// TIA Portal V20 export
FUNCTION_BLOCK "PR_StackUltraWeldSeq_Soft2"   // FB55, LAD
{ S7_Optimized_Access := 'TRUE' }
// stored: MemoryReserve 100, SetENOAutomatically false
   VAR_INPUT
      iAbort : Bool;
      iAutoRunning : Bool;
      iFaultReset : Bool;
      iPartClampClose : Bool;
      iPartClampOpen : Bool;
      iPartNotWorkable : Bool;
      iPartWorkable : Bool;
      iRFReadDone : Bool;
      iRFReadError : Bool;
      iRFWriteDone : Bool;
      iRFWriteError : Bool;
      iReject : Bool;
      iReset_fault : Bool;
      iRetry : Bool;
      iRetryCount : Int;
      iSstMode : Bool;
      iSstPB : Bool;
      iStartFrmFibroseq : Bool;
      iWeldComplete : Bool;
      iWeldTabDown : Bool;
      iWeldTabUp : Bool;
      iStartFrmFibroSeq_1 : Bool;
      iAutorunning_1 : Bool;
   END_VAR
   VAR_OUTPUT
      qError : Array[0..3] of Bool;
      qFumeExtractorON : Bool;
      qMessage : Array[0..2] of Bool;
      qPartClampClose : Bool;
      qPartClampOpen : Bool;
      qStackUltraWeldOver : Bool;
      qWeldTabDown : Bool;
      qWeldTabUp : Bool;
   END_VAR
   VAR
      c20_ChkRecovery_T1 : Bool;
      c20_ChkRecovery_T2 : Bool;
      c20_ChkRecovery_T3 : Bool;
      c21_WtRFIDReadOver_T1 : Bool;
      c21_WtRFIDReadOver_T2 : Bool;
      c22_ChkReadRetryCnt_T1 : Bool;
      c22_ChkReadRetryCnt_T2 : Bool;
      c23_ChkPartWrkSts_T1 : Bool;
      c23_ChkPartWrkSts_T2 : Bool;
      c24_WtOpDecision_T1 : Bool;
      c24_WtOpDecision_T2 : Bool;
      c81_WtRFIDWriteOver_T1 : Bool;
      c81_WtRFIDWriteOver_T2 : Bool;
      c82_ChkWriteRetryCnt_T1 : Bool;
      c82_ChkWriteRetryCnt_T2 : Bool;
      c83_WtOpDecisionWrite_T1 : Bool;
      c83_WtOpDecisionWrite_T2 : Bool;
      StateNo : Int;
      s10_WtStartFrmFibro : Bool;
      s10_WtStartFrmFibro_T1 : Bool;
      s1_WtResetRel : Bool;
      s1_WtResetRel_T1 : Bool;
      s20_ChkRecovery : Bool;
      s20_ChkRecovery_T1 : Bool;
      s20_ChkRecovery_T2 : Bool;
      s20_ChkRecovery_T3 : Bool;
      s21_WtRFIDReadOver : Bool;
      s21_WtRFIDReadOver_T1 : Bool;
      s21_WtRFIDReadOver_T2 : Bool;
      s22_ChkReadRetryCnt : Bool;
      s22_ChkReadRetryCnt_T1 : Bool;
      s22_ChkReadRetryCnt_T2 : Bool;
      s23_ChkPartWrkSts : Bool;
      s23_ChkPartWrkSts_T1 : Bool;
      s23_ChkPartWrkSts_T2 : Bool;
      s24_WtOpDecision : Bool;
      s24_WtOpDecision_T1 : Bool;
      s24_WtOpDecision_T2 : Bool;
      s30_WtOpAck : Bool;
      s30_WtOpAck_T1 : Bool;
      s40_WtPartClamp : Bool;
      s40_WtPartClamp_T1 : Bool;
      s50_WtWeldTabDown : Bool;
      s50_WtWeldTabDown_T1 : Bool;
      s60_WtWeldComplete : Bool;
      s60_WtWeldComplete_T1 : Bool;
      s70_WtWeldTabUp : Bool;
      s70_WtWeldTabUp_T1 : Bool;
      s80_WtPartClampOpen : Bool;
      s80_WtPartClampOpen_T1 : Bool;
      s81_WtRFIDWriteOver : Bool;
      s81_WtRFIDWriteOver_T1 : Bool;
      s81_WtRFIDWriteOver_T2 : Bool;
      s82_ChkWriteRetryCnt : Bool;
      s82_ChkWriteRetryCnt_T1 : Bool;
      s82_ChkWriteRetryCnt_T2 : Bool;
      s83_WtOpDecisionWrite : Bool;
      s83_WtOpDecisionWrite_T1 : Bool;
      s83_WtOpDecisionWrite_T2 : Bool;
      s90_WtStartLow : Bool;
      s90_WtStartLow_T1 : Bool;
      sRFReadRetryCount : Int;
      sRFWriteRetryCount : Int;
      sSst : Bool;
      sSstPulse : Bool;
      sSstRise : Bool;
      sStWtResetRel : Bool;
      sStWtResetRel_T1 : Bool;
      sWeldDlyOver : Bool;
      sweldingInProgress : Int;
      SET : Bool;
      c20_ChkRecovery_clamp : Bool;
   END_VAR
   VAR_TEMP
      tOne : Bool;
      tRFReadRetryCountInc : Int;
      tRFWriteRetryCountInc : Int;
   END_VAR
   VAR_TEMP   // added for the SCL form of the ladder/FBD networks
      _w1 : Bool;
      _w2 : Bool;
   END_VAR
BEGIN

REGION Network 1
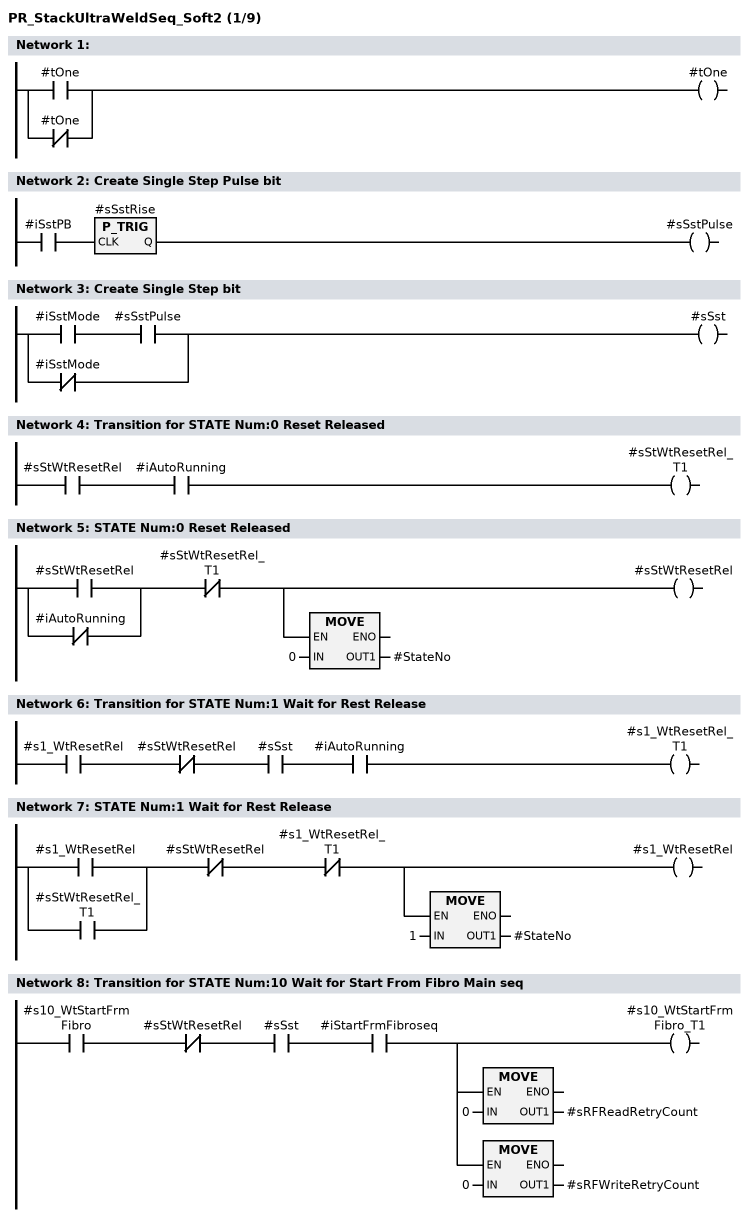
   RUNG wire#powerrail
      Contact( #tOne )
      wire#w1
      Coil( #tOne )
   END_RUNG
   RUNG wire#powerrail
      I_Contact( #tOne )
   END_RUNG wire#w1
   // the same network as SCL:
   #tOne := #tOne OR NOT #tOne;
END_REGION

REGION Network 2: Create Single Step Pulse bit
   RUNG wire#powerrail
      Contact( #iSstPB )
      P_Trig( #sSstRise )
      Coil( #sSstPulse )
   END_RUNG
   // the same network as SCL:
   #_w1 := #iSstPB AND NOT #sSstRise;   // rising edge
   #sSstRise := #iSstPB;
   #sSstPulse := #_w1;
END_REGION

REGION Network 3: Create Single Step bit
   RUNG wire#powerrail
      Contact( #iSstMode )
      Contact( #sSstPulse )
      wire#w1
      Coil( #sSst )
   END_RUNG
   RUNG wire#powerrail
      I_Contact( #iSstMode )
   END_RUNG wire#w1
   // the same network as SCL:
   #sSst := (#iSstMode AND #sSstPulse) OR NOT #iSstMode;
END_REGION

REGION Network 4: Transition for STATE Num:0 Reset Released
   RUNG wire#powerrail
      Contact( #sStWtResetRel )
      Contact( #iAutoRunning )
      Coil( #sStWtResetRel_T1 )
   END_RUNG
   // the same network as SCL:
   #sStWtResetRel_T1 := #sStWtResetRel AND #iAutoRunning;
END_REGION

REGION Network 5: STATE Num:0 Reset Released
   RUNG wire#powerrail
      Contact( #sStWtResetRel )
      wire#w1
      I_Contact( #sStWtResetRel_T1 )
      wire#w2
      Coil( #sStWtResetRel )
   END_RUNG
   RUNG wire#powerrail
      I_Contact( #iAutoRunning )
   END_RUNG wire#w1
   RUNG wire#w2
      { S7_GenerateENO := "TRUE" } Move(in := 0, out1 => #StateNo)
   END_RUNG
   // the same network as SCL:
   #sStWtResetRel := (#sStWtResetRel OR NOT #iAutoRunning) AND NOT #sStWtResetRel_T1;
   IF #sStWtResetRel THEN #StateNo := 0; END_IF;
END_REGION

REGION Network 6: Transition for STATE Num:1 Wait for Rest Release
   RUNG wire#powerrail
      Contact( #s1_WtResetRel )
      I_Contact( #sStWtResetRel )
      Contact( #sSst )
      Contact( #iAutoRunning )
      Coil( #s1_WtResetRel_T1 )
   END_RUNG
   // the same network as SCL:
   #s1_WtResetRel_T1 := #s1_WtResetRel AND NOT #sStWtResetRel AND #sSst AND #iAutoRunning;
END_REGION

REGION Network 7: STATE Num:1 Wait for Rest Release
   RUNG wire#powerrail
      Contact( #s1_WtResetRel )
      wire#w1
      I_Contact( #sStWtResetRel )
      I_Contact( #s1_WtResetRel_T1 )
      wire#w2
      Coil( #s1_WtResetRel )
   END_RUNG
   RUNG wire#powerrail
      Contact( #sStWtResetRel_T1 )
   END_RUNG wire#w1
   RUNG wire#w2
      { S7_GenerateENO := "TRUE" } Move(in := 1, out1 => #StateNo)
   END_RUNG
   // the same network as SCL:
   #s1_WtResetRel := (#s1_WtResetRel OR #sStWtResetRel_T1) AND NOT #sStWtResetRel AND NOT #s1_WtResetRel_T1;
   IF #s1_WtResetRel THEN #StateNo := 1; END_IF;
END_REGION

REGION Network 8: Transition for STATE Num:10 Wait for Start From Fibro Main seq
   RUNG wire#powerrail
      Contact( #s10_WtStartFrmFibro )
      I_Contact( #sStWtResetRel )
      Contact( #sSst )
      Contact( #iStartFrmFibroseq )
      wire#w1
      Coil( #s10_WtStartFrmFibro_T1 )
   END_RUNG
   RUNG wire#w1
      Move(in := 0, out1 => #sRFReadRetryCount)
   END_RUNG
   RUNG wire#w1
      Move(in := 0, out1 => #sRFWriteRetryCount)
   END_RUNG
   // the same network as SCL:
   #s10_WtStartFrmFibro_T1 := #s10_WtStartFrmFibro AND NOT #sStWtResetRel AND #sSst AND #iStartFrmFibroseq;
   IF #s10_WtStartFrmFibro_T1 THEN
       #sRFReadRetryCount := 0;
       #sRFWriteRetryCount := 0;
   END_IF;
END_REGION

REGION Network 9: STATE Num:10 Wait for Start From Fibro Main seq
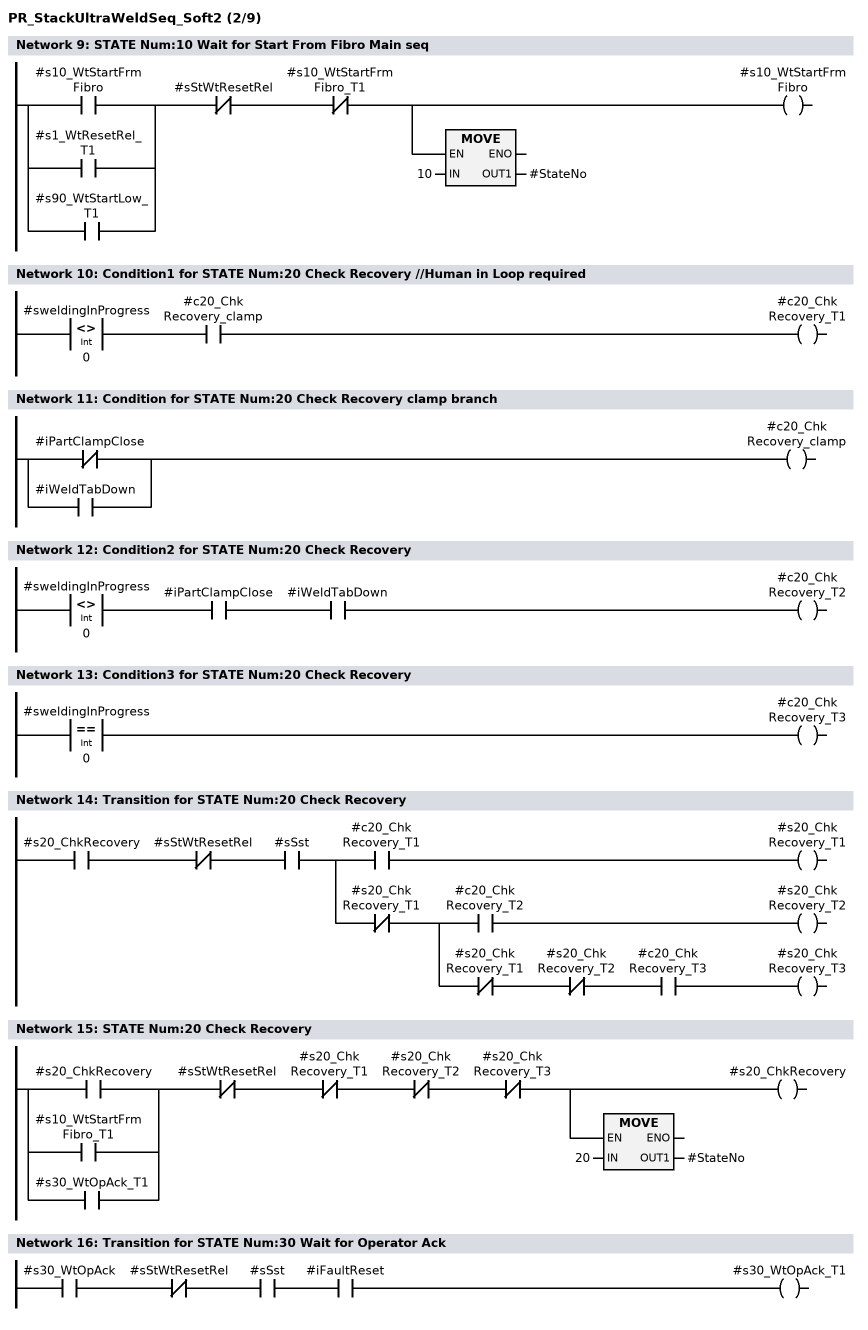
   RUNG wire#powerrail
      Contact( #s10_WtStartFrmFibro )
      wire#w1
      I_Contact( #sStWtResetRel )
      I_Contact( #s10_WtStartFrmFibro_T1 )
      wire#w2
      Coil( #s10_WtStartFrmFibro )
   END_RUNG
   RUNG wire#powerrail
      Contact( #s1_WtResetRel_T1 )
   END_RUNG wire#w1
   RUNG wire#powerrail
      Contact( #s90_WtStartLow_T1 )
   END_RUNG wire#w1
   RUNG wire#w2
      { S7_GenerateENO := "TRUE" } Move(in := 10, out1 => #StateNo)
   END_RUNG
   // the same network as SCL:
   #s10_WtStartFrmFibro := (#s10_WtStartFrmFibro OR #s1_WtResetRel_T1 OR #s90_WtStartLow_T1) AND NOT #sStWtResetRel AND NOT #s10_WtStartFrmFibro_T1;
   IF #s10_WtStartFrmFibro THEN #StateNo := 10; END_IF;
END_REGION

REGION Network 10: Condition1 for STATE Num:20 Check Recovery //Human in Loop required
   RUNG wire#powerrail
      { S7_Templates := "SrcType := Int" } NE_Contact(in1 := #sweldingInProgress, in2 := 0)
      Contact( #c20_ChkRecovery_clamp )
      Coil( #c20_ChkRecovery_T1 )
   END_RUNG
   // the same network as SCL:
   #c20_ChkRecovery_T1 := (#sweldingInProgress <> 0) AND #c20_ChkRecovery_clamp;
END_REGION

REGION Network 11: Condition for STATE Num:20 Check Recovery clamp branch
   RUNG wire#powerrail
      I_Contact( #iPartClampClose )
      wire#w1
      Coil( #c20_ChkRecovery_clamp )
   END_RUNG
   RUNG wire#powerrail
      Contact( #iWeldTabDown )
   END_RUNG wire#w1
   // the same network as SCL:
   #c20_ChkRecovery_clamp := NOT #iPartClampClose OR #iWeldTabDown;
END_REGION

REGION Network 12: Condition2 for STATE Num:20 Check Recovery
   RUNG wire#powerrail
      { S7_Templates := "SrcType := Int" } NE_Contact(in1 := #sweldingInProgress, in2 := 0)
      Contact( #iPartClampClose )
      Contact( #iWeldTabDown )
      Coil( #c20_ChkRecovery_T2 )
   END_RUNG
   // the same network as SCL:
   #c20_ChkRecovery_T2 := (#sweldingInProgress <> 0) AND #iPartClampClose AND #iWeldTabDown;
END_REGION

REGION Network 13: Condition3 for STATE Num:20 Check Recovery
   RUNG wire#powerrail
      { S7_Templates := "SrcType := Int" } EQ_Contact(in1 := #sweldingInProgress, in2 := 0)
      Coil( #c20_ChkRecovery_T3 )
   END_RUNG
   // the same network as SCL:
   #c20_ChkRecovery_T3 := #sweldingInProgress = 0;
END_REGION

REGION Network 14: Transition for STATE Num:20 Check Recovery
   RUNG wire#powerrail
      Contact( #s20_ChkRecovery )
      I_Contact( #sStWtResetRel )
      Contact( #sSst )
      wire#w1
      Contact( #c20_ChkRecovery_T1 )
      Coil( #s20_ChkRecovery_T1 )
   END_RUNG
   RUNG wire#w1
      I_Contact( #s20_ChkRecovery_T1 )
      wire#w2
      Contact( #c20_ChkRecovery_T2 )
      Coil( #s20_ChkRecovery_T2 )
   END_RUNG
   RUNG wire#w2
      I_Contact( #s20_ChkRecovery_T1 )
      I_Contact( #s20_ChkRecovery_T2 )
      Contact( #c20_ChkRecovery_T3 )
      Coil( #s20_ChkRecovery_T3 )
   END_RUNG
   // the same network as SCL:
   #_w1 := #s20_ChkRecovery AND NOT #sStWtResetRel AND #sSst;
   #s20_ChkRecovery_T1 := #_w1 AND #c20_ChkRecovery_T1;
   #_w2 := #_w1 AND NOT #s20_ChkRecovery_T1;
   #s20_ChkRecovery_T2 := #_w2 AND #c20_ChkRecovery_T2;
   #s20_ChkRecovery_T3 := #_w2 AND NOT #s20_ChkRecovery_T1 AND NOT #s20_ChkRecovery_T2 AND #c20_ChkRecovery_T3;
END_REGION

REGION Network 15: STATE Num:20 Check Recovery
   RUNG wire#powerrail
      Contact( #s20_ChkRecovery )
      wire#w1
      I_Contact( #sStWtResetRel )
      I_Contact( #s20_ChkRecovery_T1 )
      I_Contact( #s20_ChkRecovery_T2 )
      I_Contact( #s20_ChkRecovery_T3 )
      wire#w2
      Coil( #s20_ChkRecovery )
   END_RUNG
   RUNG wire#powerrail
      Contact( #s10_WtStartFrmFibro_T1 )
   END_RUNG wire#w1
   RUNG wire#powerrail
      Contact( #s30_WtOpAck_T1 )
   END_RUNG wire#w1
   RUNG wire#w2
      { S7_GenerateENO := "TRUE" } Move(in := 20, out1 => #StateNo)
   END_RUNG
   // the same network as SCL:
   #s20_ChkRecovery := (#s20_ChkRecovery OR #s10_WtStartFrmFibro_T1 OR #s30_WtOpAck_T1) AND NOT #sStWtResetRel AND NOT #s20_ChkRecovery_T1 AND NOT #s20_ChkRecovery_T2 AND NOT #s20_ChkRecovery_T3;
   IF #s20_ChkRecovery THEN #StateNo := 20; END_IF;
END_REGION

REGION Network 16: Transition for STATE Num:30 Wait for Operator Ack
   RUNG wire#powerrail
      Contact( #s30_WtOpAck )
      I_Contact( #sStWtResetRel )
      Contact( #sSst )
      Contact( #iFaultReset )
      Coil( #s30_WtOpAck_T1 )
   END_RUNG
   // the same network as SCL:
   #s30_WtOpAck_T1 := #s30_WtOpAck AND NOT #sStWtResetRel AND #sSst AND #iFaultReset;
END_REGION

REGION Network 17: STATE Num:30 Wait for Operator Ack
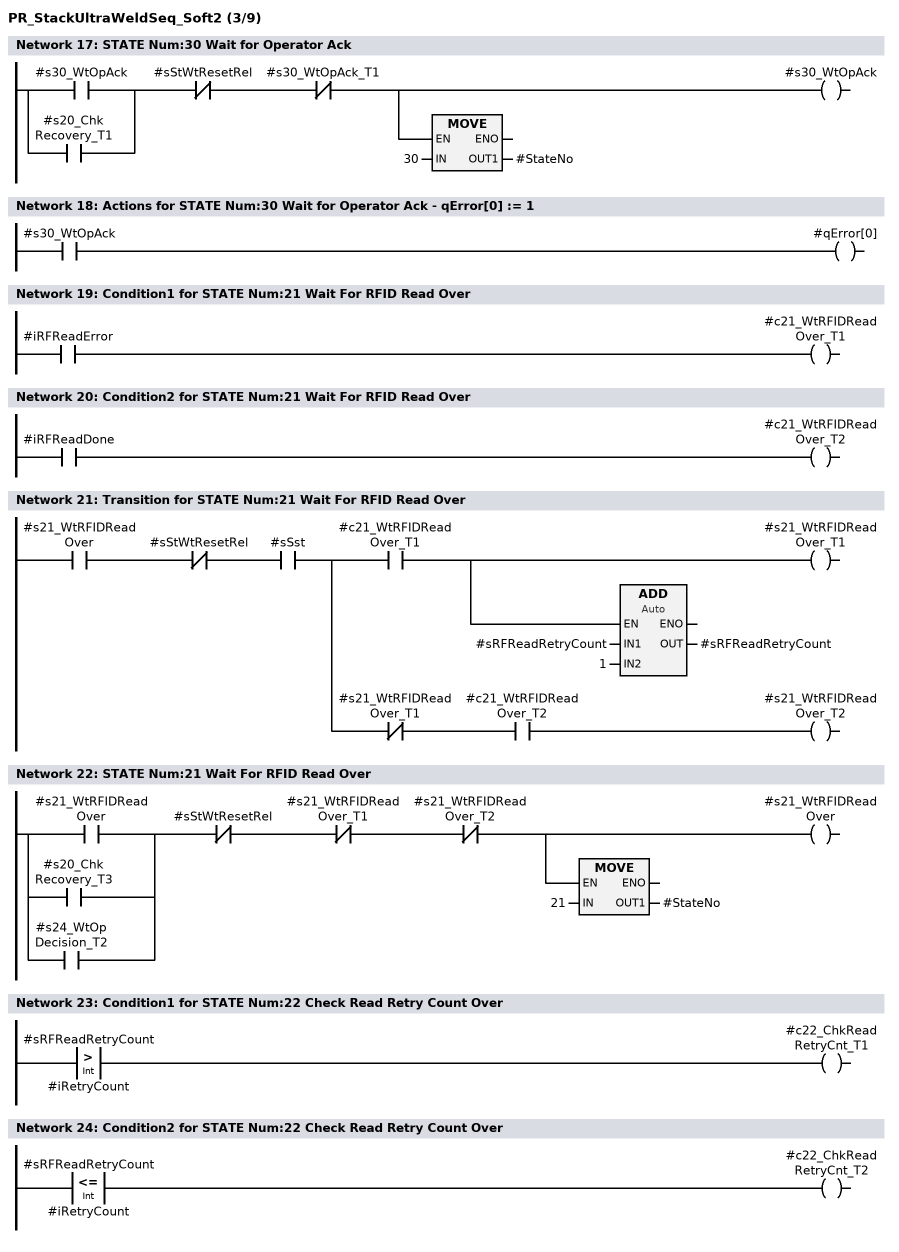
   RUNG wire#powerrail
      Contact( #s30_WtOpAck )
      wire#w1
      I_Contact( #sStWtResetRel )
      I_Contact( #s30_WtOpAck_T1 )
      wire#w2
      Coil( #s30_WtOpAck )
   END_RUNG
   RUNG wire#powerrail
      Contact( #s20_ChkRecovery_T1 )
   END_RUNG wire#w1
   RUNG wire#w2
      { S7_GenerateENO := "TRUE" } Move(in := 30, out1 => #StateNo)
   END_RUNG
   // the same network as SCL:
   #s30_WtOpAck := (#s30_WtOpAck OR #s20_ChkRecovery_T1) AND NOT #sStWtResetRel AND NOT #s30_WtOpAck_T1;
   IF #s30_WtOpAck THEN #StateNo := 30; END_IF;
END_REGION

REGION Network 18: Actions for STATE Num:30 Wait for Operator Ack - qError[0] := 1
   RUNG wire#powerrail
      Contact( #s30_WtOpAck )
      Coil( #qError[0] )
   END_RUNG
   // the same network as SCL:
   #qError[0] := #s30_WtOpAck;
END_REGION

REGION Network 19: Condition1 for STATE Num:21 Wait For RFID Read Over
   RUNG wire#powerrail
      Contact( #iRFReadError )
      Coil( #c21_WtRFIDReadOver_T1 )
   END_RUNG
   // the same network as SCL:
   #c21_WtRFIDReadOver_T1 := #iRFReadError;
END_REGION

REGION Network 20: Condition2 for STATE Num:21 Wait For RFID Read Over
   RUNG wire#powerrail
      Contact( #iRFReadDone )
      Coil( #c21_WtRFIDReadOver_T2 )
   END_RUNG
   // the same network as SCL:
   #c21_WtRFIDReadOver_T2 := #iRFReadDone;
END_REGION

REGION Network 21: Transition for STATE Num:21 Wait For RFID Read Over
   RUNG wire#powerrail
      Contact( #s21_WtRFIDReadOver )
      I_Contact( #sStWtResetRel )
      Contact( #sSst )
      wire#w1
      Contact( #c21_WtRFIDReadOver_T1 )
      wire#w2
      Coil( #s21_WtRFIDReadOver_T1 )
   END_RUNG
   RUNG wire#w2
      Add(in1 := #sRFReadRetryCount, in2 := 1, out => #sRFReadRetryCount)
   END_RUNG
   RUNG wire#w1
      I_Contact( #s21_WtRFIDReadOver_T1 )
      Contact( #c21_WtRFIDReadOver_T2 )
      Coil( #s21_WtRFIDReadOver_T2 )
   END_RUNG
   // the same network as SCL:
   #_w1 := #s21_WtRFIDReadOver AND NOT #sStWtResetRel AND #sSst;
   #s21_WtRFIDReadOver_T1 := #_w1 AND #c21_WtRFIDReadOver_T1;
   IF #s21_WtRFIDReadOver_T1 THEN #sRFReadRetryCount := #sRFReadRetryCount + 1; END_IF;
   #s21_WtRFIDReadOver_T2 := #_w1 AND NOT #s21_WtRFIDReadOver_T1 AND #c21_WtRFIDReadOver_T2;
END_REGION

REGION Network 22: STATE Num:21 Wait For RFID Read Over
   RUNG wire#powerrail
      Contact( #s21_WtRFIDReadOver )
      wire#w1
      I_Contact( #sStWtResetRel )
      I_Contact( #s21_WtRFIDReadOver_T1 )
      I_Contact( #s21_WtRFIDReadOver_T2 )
      wire#w2
      Coil( #s21_WtRFIDReadOver )
   END_RUNG
   RUNG wire#powerrail
      Contact( #s20_ChkRecovery_T3 )
   END_RUNG wire#w1
   RUNG wire#powerrail
      Contact( #s24_WtOpDecision_T2 )
   END_RUNG wire#w1
   RUNG wire#w2
      { S7_GenerateENO := "TRUE" } Move(in := 21, out1 => #StateNo)
   END_RUNG
   // the same network as SCL:
   #s21_WtRFIDReadOver := (#s21_WtRFIDReadOver OR #s20_ChkRecovery_T3 OR #s24_WtOpDecision_T2) AND NOT #sStWtResetRel AND NOT #s21_WtRFIDReadOver_T1 AND NOT #s21_WtRFIDReadOver_T2;
   IF #s21_WtRFIDReadOver THEN #StateNo := 21; END_IF;
END_REGION

REGION Network 23: Condition1 for STATE Num:22 Check Read Retry Count Over
   RUNG wire#powerrail
      { S7_Templates := "SrcType := Int" } GT_Contact(in1 := #sRFReadRetryCount, in2 := #iRetryCount)
      Coil( #c22_ChkReadRetryCnt_T1 )
   END_RUNG
   // the same network as SCL:
   #c22_ChkReadRetryCnt_T1 := #sRFReadRetryCount > #iRetryCount;
END_REGION

REGION Network 24: Condition2 for STATE Num:22 Check Read Retry Count Over
   RUNG wire#powerrail
      { S7_Templates := "SrcType := Int" } LE_Contact(in1 := #sRFReadRetryCount, in2 := #iRetryCount)
      Coil( #c22_ChkReadRetryCnt_T2 )
   END_RUNG
   // the same network as SCL:
   #c22_ChkReadRetryCnt_T2 := #sRFReadRetryCount <= #iRetryCount;
END_REGION

REGION Network 25: Transition for STATE Num:22 Check Read Retry Count Over
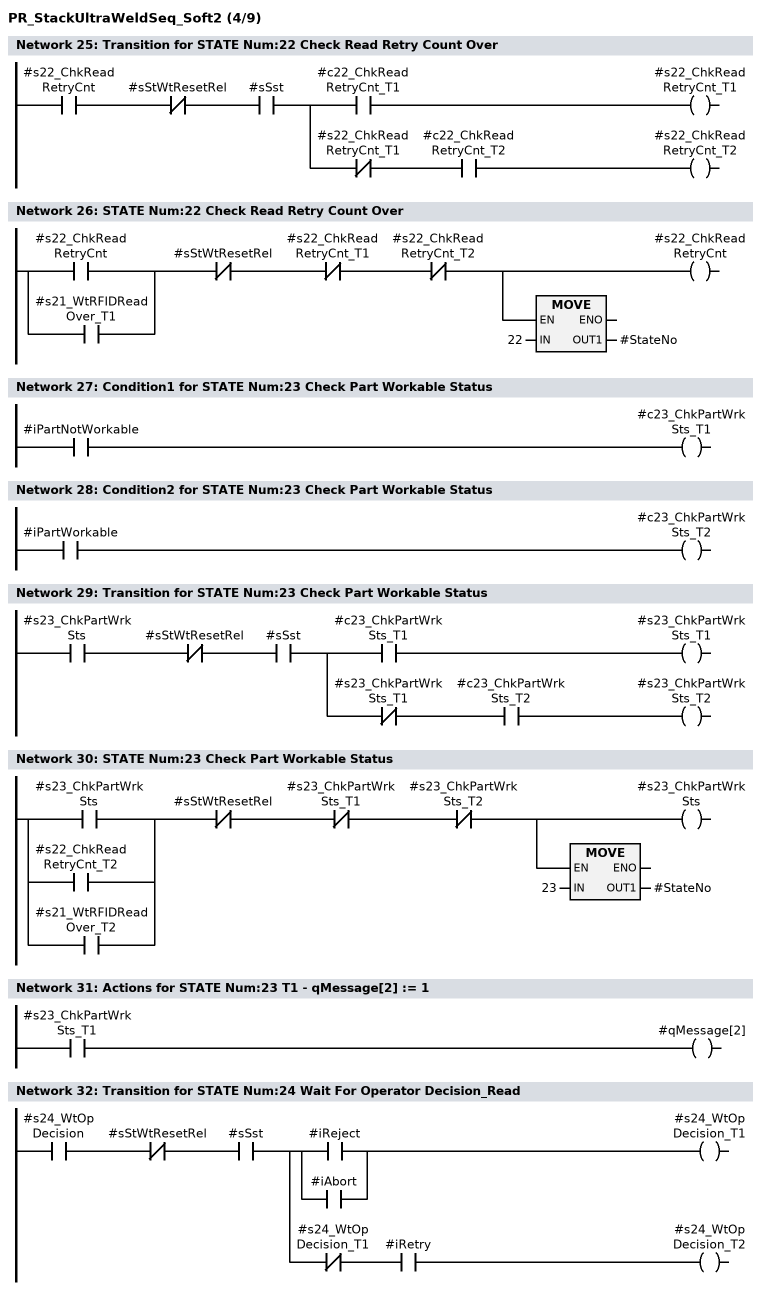
   RUNG wire#powerrail
      Contact( #s22_ChkReadRetryCnt )
      I_Contact( #sStWtResetRel )
      Contact( #sSst )
      wire#w1
      Contact( #c22_ChkReadRetryCnt_T1 )
      Coil( #s22_ChkReadRetryCnt_T1 )
   END_RUNG
   RUNG wire#w1
      I_Contact( #s22_ChkReadRetryCnt_T1 )
      Contact( #c22_ChkReadRetryCnt_T2 )
      Coil( #s22_ChkReadRetryCnt_T2 )
   END_RUNG
   // the same network as SCL:
   #_w1 := #s22_ChkReadRetryCnt AND NOT #sStWtResetRel AND #sSst;
   #s22_ChkReadRetryCnt_T1 := #_w1 AND #c22_ChkReadRetryCnt_T1;
   #s22_ChkReadRetryCnt_T2 := #_w1 AND NOT #s22_ChkReadRetryCnt_T1 AND #c22_ChkReadRetryCnt_T2;
END_REGION

REGION Network 26: STATE Num:22 Check Read Retry Count Over
   RUNG wire#powerrail
      Contact( #s22_ChkReadRetryCnt )
      wire#w1
      I_Contact( #sStWtResetRel )
      I_Contact( #s22_ChkReadRetryCnt_T1 )
      I_Contact( #s22_ChkReadRetryCnt_T2 )
      wire#w2
      Coil( #s22_ChkReadRetryCnt )
   END_RUNG
   RUNG wire#powerrail
      Contact( #s21_WtRFIDReadOver_T1 )
   END_RUNG wire#w1
   RUNG wire#w2
      { S7_GenerateENO := "TRUE" } Move(in := 22, out1 => #StateNo)
   END_RUNG
   // the same network as SCL:
   #s22_ChkReadRetryCnt := (#s22_ChkReadRetryCnt OR #s21_WtRFIDReadOver_T1) AND NOT #sStWtResetRel AND NOT #s22_ChkReadRetryCnt_T1 AND NOT #s22_ChkReadRetryCnt_T2;
   IF #s22_ChkReadRetryCnt THEN #StateNo := 22; END_IF;
END_REGION

REGION Network 27: Condition1 for STATE Num:23 Check Part Workable Status
   RUNG wire#powerrail
      Contact( #iPartNotWorkable )
      Coil( #c23_ChkPartWrkSts_T1 )
   END_RUNG
   // the same network as SCL:
   #c23_ChkPartWrkSts_T1 := #iPartNotWorkable;
END_REGION

REGION Network 28: Condition2 for STATE Num:23 Check Part Workable Status
   RUNG wire#powerrail
      Contact( #iPartWorkable )
      Coil( #c23_ChkPartWrkSts_T2 )
   END_RUNG
   // the same network as SCL:
   #c23_ChkPartWrkSts_T2 := #iPartWorkable;
END_REGION

REGION Network 29: Transition for STATE Num:23 Check Part Workable Status
   RUNG wire#powerrail
      Contact( #s23_ChkPartWrkSts )
      I_Contact( #sStWtResetRel )
      Contact( #sSst )
      wire#w1
      Contact( #c23_ChkPartWrkSts_T1 )
      Coil( #s23_ChkPartWrkSts_T1 )
   END_RUNG
   RUNG wire#w1
      I_Contact( #s23_ChkPartWrkSts_T1 )
      Contact( #c23_ChkPartWrkSts_T2 )
      Coil( #s23_ChkPartWrkSts_T2 )
   END_RUNG
   // the same network as SCL:
   #_w1 := #s23_ChkPartWrkSts AND NOT #sStWtResetRel AND #sSst;
   #s23_ChkPartWrkSts_T1 := #_w1 AND #c23_ChkPartWrkSts_T1;
   #s23_ChkPartWrkSts_T2 := #_w1 AND NOT #s23_ChkPartWrkSts_T1 AND #c23_ChkPartWrkSts_T2;
END_REGION

REGION Network 30: STATE Num:23 Check Part Workable Status
   RUNG wire#powerrail
      Contact( #s23_ChkPartWrkSts )
      wire#w1
      I_Contact( #sStWtResetRel )
      I_Contact( #s23_ChkPartWrkSts_T1 )
      I_Contact( #s23_ChkPartWrkSts_T2 )
      wire#w2
      Coil( #s23_ChkPartWrkSts )
   END_RUNG
   RUNG wire#powerrail
      Contact( #s22_ChkReadRetryCnt_T2 )
   END_RUNG wire#w1
   RUNG wire#powerrail
      Contact( #s21_WtRFIDReadOver_T2 )
   END_RUNG wire#w1
   RUNG wire#w2
      { S7_GenerateENO := "TRUE" } Move(in := 23, out1 => #StateNo)
   END_RUNG
   // the same network as SCL:
   #s23_ChkPartWrkSts := (#s23_ChkPartWrkSts OR #s22_ChkReadRetryCnt_T2 OR #s21_WtRFIDReadOver_T2) AND NOT #sStWtResetRel AND NOT #s23_ChkPartWrkSts_T1 AND NOT #s23_ChkPartWrkSts_T2;
   IF #s23_ChkPartWrkSts THEN #StateNo := 23; END_IF;
END_REGION

REGION Network 31: Actions for STATE Num:23 T1 - qMessage[2] := 1
   RUNG wire#powerrail
      Contact( #s23_ChkPartWrkSts_T1 )
      Coil( #qMessage[2] )
   END_RUNG
   // the same network as SCL:
   #qMessage[2] := #s23_ChkPartWrkSts_T1;
END_REGION

REGION Network 32: Transition for STATE Num:24 Wait For Operator Decision_Read
   RUNG wire#powerrail
      Contact( #s24_WtOpDecision )
      I_Contact( #sStWtResetRel )
      Contact( #sSst )
      wire#w1
      Contact( #iReject )
      wire#w2
      Coil( #s24_WtOpDecision_T1 )
   END_RUNG
   RUNG wire#w1
      Contact( #iAbort )
   END_RUNG wire#w2
   RUNG wire#w1
      I_Contact( #s24_WtOpDecision_T1 )
      Contact( #iRetry )
      Coil( #s24_WtOpDecision_T2 )
   END_RUNG
   // the same network as SCL:
   #_w1 := #s24_WtOpDecision AND NOT #sStWtResetRel AND #sSst;
   #s24_WtOpDecision_T1 := #_w1 AND (#iReject OR #iAbort);
   #s24_WtOpDecision_T2 := #_w1 AND NOT #s24_WtOpDecision_T1 AND #iRetry;
END_REGION

REGION Network 33: STATE Num:24 Wait For Operator Decision_Read
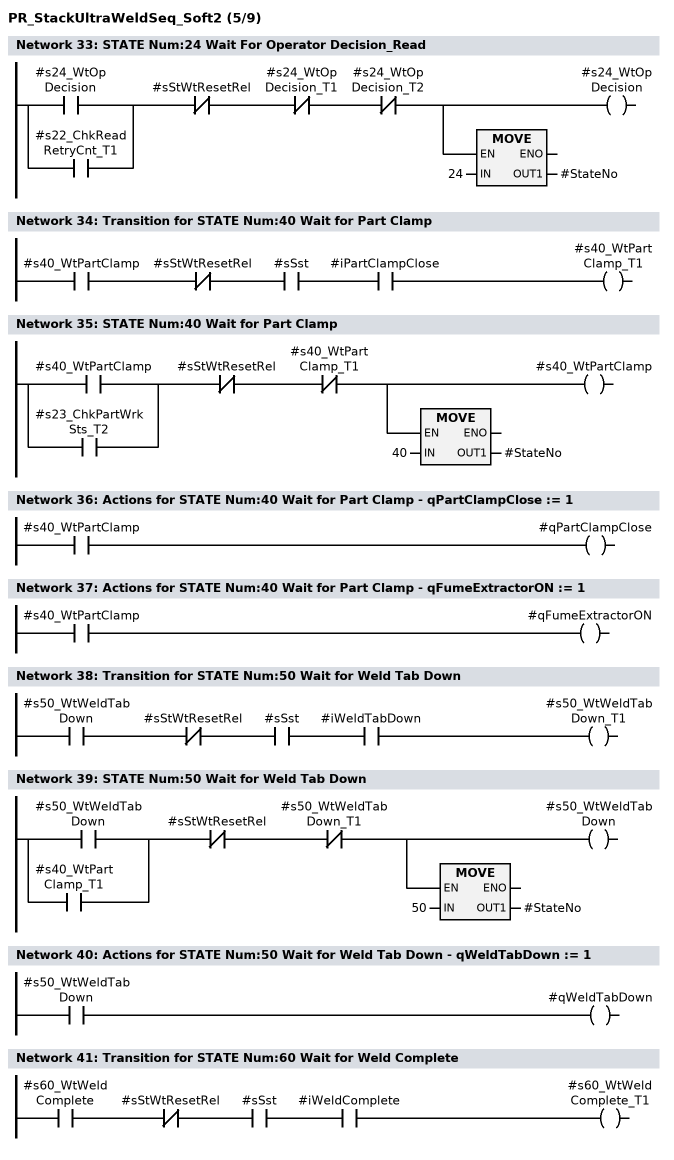
   RUNG wire#powerrail
      Contact( #s24_WtOpDecision )
      wire#w1
      I_Contact( #sStWtResetRel )
      I_Contact( #s24_WtOpDecision_T1 )
      I_Contact( #s24_WtOpDecision_T2 )
      wire#w2
      Coil( #s24_WtOpDecision )
   END_RUNG
   RUNG wire#powerrail
      Contact( #s22_ChkReadRetryCnt_T1 )
   END_RUNG wire#w1
   RUNG wire#w2
      { S7_GenerateENO := "TRUE" } Move(in := 24, out1 => #StateNo)
   END_RUNG
   // the same network as SCL:
   #s24_WtOpDecision := (#s24_WtOpDecision OR #s22_ChkReadRetryCnt_T1) AND NOT #sStWtResetRel AND NOT #s24_WtOpDecision_T1 AND NOT #s24_WtOpDecision_T2;
   IF #s24_WtOpDecision THEN #StateNo := 24; END_IF;
END_REGION

REGION Network 34: Transition for STATE Num:40 Wait for Part Clamp
   RUNG wire#powerrail
      Contact( #s40_WtPartClamp )
      I_Contact( #sStWtResetRel )
      Contact( #sSst )
      Contact( #iPartClampClose )
      Coil( #s40_WtPartClamp_T1 )
   END_RUNG
   // the same network as SCL:
   #s40_WtPartClamp_T1 := #s40_WtPartClamp AND NOT #sStWtResetRel AND #sSst AND #iPartClampClose;
END_REGION

REGION Network 35: STATE Num:40 Wait for Part Clamp
   RUNG wire#powerrail
      Contact( #s40_WtPartClamp )
      wire#w1
      I_Contact( #sStWtResetRel )
      I_Contact( #s40_WtPartClamp_T1 )
      wire#w2
      Coil( #s40_WtPartClamp )
   END_RUNG
   RUNG wire#powerrail
      Contact( #s23_ChkPartWrkSts_T2 )
   END_RUNG wire#w1
   RUNG wire#w2
      { S7_GenerateENO := "TRUE" } Move(in := 40, out1 => #StateNo)
   END_RUNG
   // the same network as SCL:
   #s40_WtPartClamp := (#s40_WtPartClamp OR #s23_ChkPartWrkSts_T2) AND NOT #sStWtResetRel AND NOT #s40_WtPartClamp_T1;
   IF #s40_WtPartClamp THEN #StateNo := 40; END_IF;
END_REGION

REGION Network 36: Actions for STATE Num:40 Wait for Part Clamp - qPartClampClose := 1
   RUNG wire#powerrail
      Contact( #s40_WtPartClamp )
      Coil( #qPartClampClose )
   END_RUNG
   // the same network as SCL:
   #qPartClampClose := #s40_WtPartClamp;
END_REGION

REGION Network 37: Actions for STATE Num:40 Wait for Part Clamp - qFumeExtractorON := 1
   RUNG wire#powerrail
      Contact( #s40_WtPartClamp )
      Coil( #qFumeExtractorON )
   END_RUNG
   // the same network as SCL:
   #qFumeExtractorON := #s40_WtPartClamp;
END_REGION

REGION Network 38: Transition for STATE Num:50 Wait for Weld Tab Down
   RUNG wire#powerrail
      Contact( #s50_WtWeldTabDown )
      I_Contact( #sStWtResetRel )
      Contact( #sSst )
      Contact( #iWeldTabDown )
      Coil( #s50_WtWeldTabDown_T1 )
   END_RUNG
   // the same network as SCL:
   #s50_WtWeldTabDown_T1 := #s50_WtWeldTabDown AND NOT #sStWtResetRel AND #sSst AND #iWeldTabDown;
END_REGION

REGION Network 39: STATE Num:50 Wait for Weld Tab Down
   RUNG wire#powerrail
      Contact( #s50_WtWeldTabDown )
      wire#w1
      I_Contact( #sStWtResetRel )
      I_Contact( #s50_WtWeldTabDown_T1 )
      wire#w2
      Coil( #s50_WtWeldTabDown )
   END_RUNG
   RUNG wire#powerrail
      Contact( #s40_WtPartClamp_T1 )
   END_RUNG wire#w1
   RUNG wire#w2
      { S7_GenerateENO := "TRUE" } Move(in := 50, out1 => #StateNo)
   END_RUNG
   // the same network as SCL:
   #s50_WtWeldTabDown := (#s50_WtWeldTabDown OR #s40_WtPartClamp_T1) AND NOT #sStWtResetRel AND NOT #s50_WtWeldTabDown_T1;
   IF #s50_WtWeldTabDown THEN #StateNo := 50; END_IF;
END_REGION

REGION Network 40: Actions for STATE Num:50 Wait for Weld Tab Down - qWeldTabDown := 1
   RUNG wire#powerrail
      Contact( #s50_WtWeldTabDown )
      Coil( #qWeldTabDown )
   END_RUNG
   // the same network as SCL:
   #qWeldTabDown := #s50_WtWeldTabDown;
END_REGION

REGION Network 41: Transition for STATE Num:60 Wait for Weld Complete
   RUNG wire#powerrail
      Contact( #s60_WtWeldComplete )
      I_Contact( #sStWtResetRel )
      Contact( #sSst )
      Contact( #iWeldComplete )
      Coil( #s60_WtWeldComplete_T1 )
   END_RUNG
   // the same network as SCL:
   #s60_WtWeldComplete_T1 := #s60_WtWeldComplete AND NOT #sStWtResetRel AND #sSst AND #iWeldComplete;
END_REGION

REGION Network 42: STATE Num:60 Wait for Weld Complete
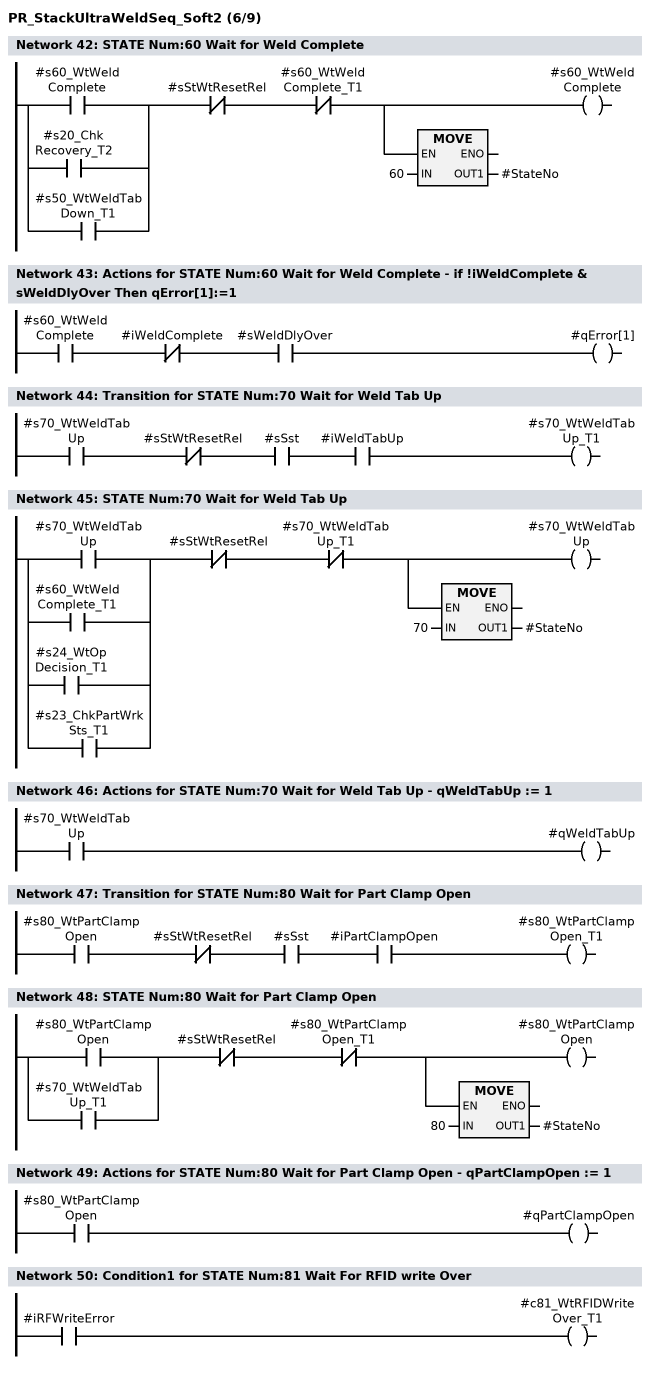
   RUNG wire#powerrail
      Contact( #s60_WtWeldComplete )
      wire#w1
      I_Contact( #sStWtResetRel )
      I_Contact( #s60_WtWeldComplete_T1 )
      wire#w2
      Coil( #s60_WtWeldComplete )
   END_RUNG
   RUNG wire#powerrail
      Contact( #s20_ChkRecovery_T2 )
   END_RUNG wire#w1
   RUNG wire#powerrail
      Contact( #s50_WtWeldTabDown_T1 )
   END_RUNG wire#w1
   RUNG wire#w2
      { S7_GenerateENO := "TRUE" } Move(in := 60, out1 => #StateNo)
   END_RUNG
   // the same network as SCL:
   #s60_WtWeldComplete := (#s60_WtWeldComplete OR #s20_ChkRecovery_T2 OR #s50_WtWeldTabDown_T1) AND NOT #sStWtResetRel AND NOT #s60_WtWeldComplete_T1;
   IF #s60_WtWeldComplete THEN #StateNo := 60; END_IF;
END_REGION

REGION Network 43: Actions for STATE Num:60 Wait for Weld Complete - if !iWeldComplete & sWeldDlyOver Then qError[1]:=1
   RUNG wire#powerrail
      Contact( #s60_WtWeldComplete )
      I_Contact( #iWeldComplete )
      Contact( #sWeldDlyOver )
      Coil( #qError[1] )
   END_RUNG
   // the same network as SCL:
   #qError[1] := #s60_WtWeldComplete AND NOT #iWeldComplete AND #sWeldDlyOver;
END_REGION

REGION Network 44: Transition for STATE Num:70 Wait for Weld Tab Up
   RUNG wire#powerrail
      Contact( #s70_WtWeldTabUp )
      I_Contact( #sStWtResetRel )
      Contact( #sSst )
      Contact( #iWeldTabUp )
      Coil( #s70_WtWeldTabUp_T1 )
   END_RUNG
   // the same network as SCL:
   #s70_WtWeldTabUp_T1 := #s70_WtWeldTabUp AND NOT #sStWtResetRel AND #sSst AND #iWeldTabUp;
END_REGION

REGION Network 45: STATE Num:70 Wait for Weld Tab Up
   RUNG wire#powerrail
      Contact( #s70_WtWeldTabUp )
      wire#w1
      I_Contact( #sStWtResetRel )
      I_Contact( #s70_WtWeldTabUp_T1 )
      wire#w2
      Coil( #s70_WtWeldTabUp )
   END_RUNG
   RUNG wire#powerrail
      Contact( #s60_WtWeldComplete_T1 )
   END_RUNG wire#w1
   RUNG wire#powerrail
      Contact( #s24_WtOpDecision_T1 )
   END_RUNG wire#w1
   RUNG wire#powerrail
      Contact( #s23_ChkPartWrkSts_T1 )
   END_RUNG wire#w1
   RUNG wire#w2
      { S7_GenerateENO := "TRUE" } Move(in := 70, out1 => #StateNo)
   END_RUNG
   // the same network as SCL:
   #s70_WtWeldTabUp := (#s70_WtWeldTabUp OR #s60_WtWeldComplete_T1 OR #s24_WtOpDecision_T1 OR #s23_ChkPartWrkSts_T1) AND NOT #sStWtResetRel AND NOT #s70_WtWeldTabUp_T1;
   IF #s70_WtWeldTabUp THEN #StateNo := 70; END_IF;
END_REGION

REGION Network 46: Actions for STATE Num:70 Wait for Weld Tab Up - qWeldTabUp := 1
   RUNG wire#powerrail
      Contact( #s70_WtWeldTabUp )
      Coil( #qWeldTabUp )
   END_RUNG
   // the same network as SCL:
   #qWeldTabUp := #s70_WtWeldTabUp;
END_REGION

REGION Network 47: Transition for STATE Num:80 Wait for Part Clamp Open
   RUNG wire#powerrail
      Contact( #s80_WtPartClampOpen )
      I_Contact( #sStWtResetRel )
      Contact( #sSst )
      Contact( #iPartClampOpen )
      Coil( #s80_WtPartClampOpen_T1 )
   END_RUNG
   // the same network as SCL:
   #s80_WtPartClampOpen_T1 := #s80_WtPartClampOpen AND NOT #sStWtResetRel AND #sSst AND #iPartClampOpen;
END_REGION

REGION Network 48: STATE Num:80 Wait for Part Clamp Open
   RUNG wire#powerrail
      Contact( #s80_WtPartClampOpen )
      wire#w1
      I_Contact( #sStWtResetRel )
      I_Contact( #s80_WtPartClampOpen_T1 )
      wire#w2
      Coil( #s80_WtPartClampOpen )
   END_RUNG
   RUNG wire#powerrail
      Contact( #s70_WtWeldTabUp_T1 )
   END_RUNG wire#w1
   RUNG wire#w2
      { S7_GenerateENO := "TRUE" } Move(in := 80, out1 => #StateNo)
   END_RUNG
   // the same network as SCL:
   #s80_WtPartClampOpen := (#s80_WtPartClampOpen OR #s70_WtWeldTabUp_T1) AND NOT #sStWtResetRel AND NOT #s80_WtPartClampOpen_T1;
   IF #s80_WtPartClampOpen THEN #StateNo := 80; END_IF;
END_REGION

REGION Network 49: Actions for STATE Num:80 Wait for Part Clamp Open - qPartClampOpen := 1
   RUNG wire#powerrail
      Contact( #s80_WtPartClampOpen )
      Coil( #qPartClampOpen )
   END_RUNG
   // the same network as SCL:
   #qPartClampOpen := #s80_WtPartClampOpen;
END_REGION

REGION Network 50: Condition1 for STATE Num:81 Wait For RFID write Over
   RUNG wire#powerrail
      Contact( #iRFWriteError )
      Coil( #c81_WtRFIDWriteOver_T1 )
   END_RUNG
   // the same network as SCL:
   #c81_WtRFIDWriteOver_T1 := #iRFWriteError;
END_REGION

REGION Network 51: Condition2 for STATE Num:81 Wait For RFID write Over
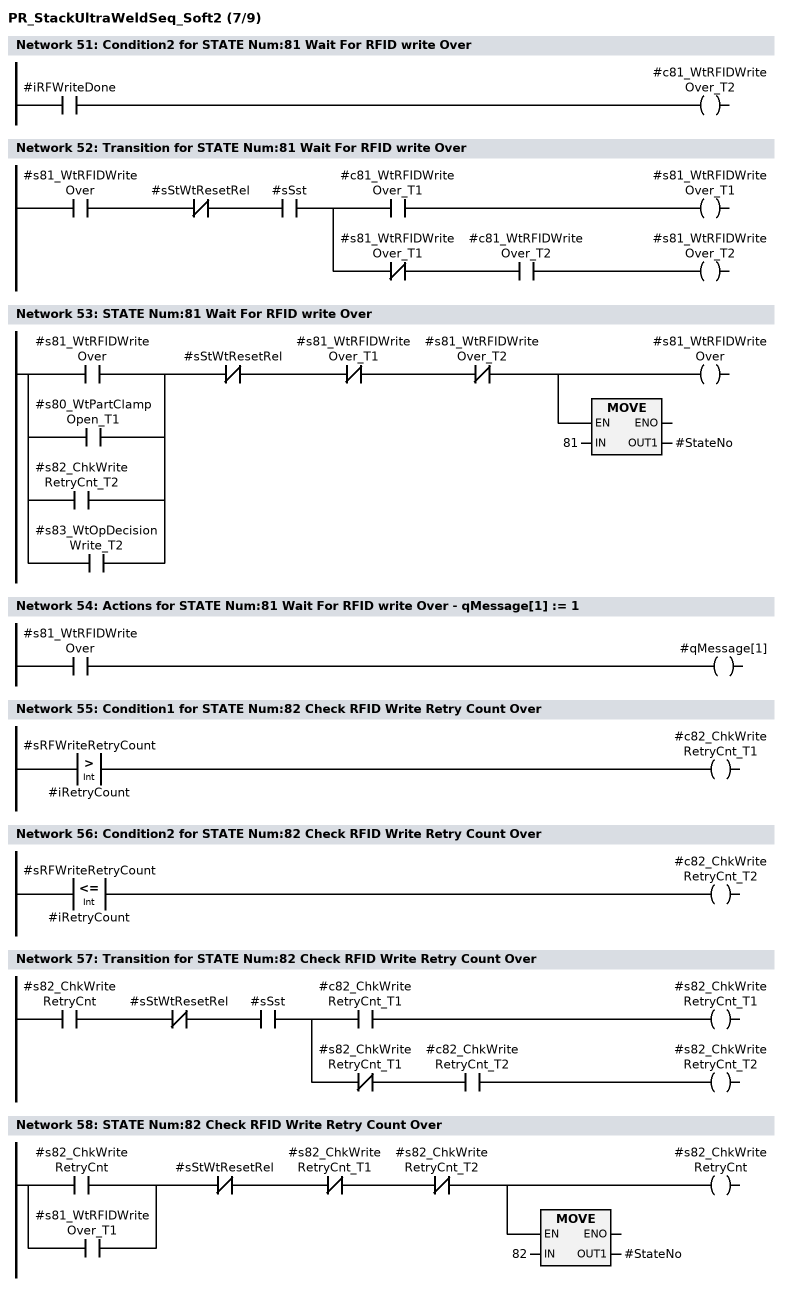
   RUNG wire#powerrail
      Contact( #iRFWriteDone )
      Coil( #c81_WtRFIDWriteOver_T2 )
   END_RUNG
   // the same network as SCL:
   #c81_WtRFIDWriteOver_T2 := #iRFWriteDone;
END_REGION

REGION Network 52: Transition for STATE Num:81 Wait For RFID write Over
   RUNG wire#powerrail
      Contact( #s81_WtRFIDWriteOver )
      I_Contact( #sStWtResetRel )
      Contact( #sSst )
      wire#w1
      Contact( #c81_WtRFIDWriteOver_T1 )
      Coil( #s81_WtRFIDWriteOver_T1 )
   END_RUNG
   RUNG wire#w1
      I_Contact( #s81_WtRFIDWriteOver_T1 )
      Contact( #c81_WtRFIDWriteOver_T2 )
      Coil( #s81_WtRFIDWriteOver_T2 )
   END_RUNG
   // the same network as SCL:
   #_w1 := #s81_WtRFIDWriteOver AND NOT #sStWtResetRel AND #sSst;
   #s81_WtRFIDWriteOver_T1 := #_w1 AND #c81_WtRFIDWriteOver_T1;
   #s81_WtRFIDWriteOver_T2 := #_w1 AND NOT #s81_WtRFIDWriteOver_T1 AND #c81_WtRFIDWriteOver_T2;
END_REGION

REGION Network 53: STATE Num:81 Wait For RFID write Over
   RUNG wire#powerrail
      Contact( #s81_WtRFIDWriteOver )
      wire#w1
      I_Contact( #sStWtResetRel )
      I_Contact( #s81_WtRFIDWriteOver_T1 )
      I_Contact( #s81_WtRFIDWriteOver_T2 )
      wire#w2
      Coil( #s81_WtRFIDWriteOver )
   END_RUNG
   RUNG wire#powerrail
      Contact( #s80_WtPartClampOpen_T1 )
   END_RUNG wire#w1
   RUNG wire#powerrail
      Contact( #s82_ChkWriteRetryCnt_T2 )
   END_RUNG wire#w1
   RUNG wire#powerrail
      Contact( #s83_WtOpDecisionWrite_T2 )
   END_RUNG wire#w1
   RUNG wire#w2
      { S7_GenerateENO := "TRUE" } Move(in := 81, out1 => #StateNo)
   END_RUNG
   // the same network as SCL:
   #s81_WtRFIDWriteOver := (#s81_WtRFIDWriteOver OR #s80_WtPartClampOpen_T1 OR #s82_ChkWriteRetryCnt_T2 OR #s83_WtOpDecisionWrite_T2) AND NOT #sStWtResetRel AND NOT #s81_WtRFIDWriteOver_T1 AND NOT #s81_WtRFIDWriteOver_T2;
   IF #s81_WtRFIDWriteOver THEN #StateNo := 81; END_IF;
END_REGION

REGION Network 54: Actions for STATE Num:81 Wait For RFID write Over - qMessage[1] := 1
   RUNG wire#powerrail
      Contact( #s81_WtRFIDWriteOver )
      Coil( #qMessage[1] )
   END_RUNG
   // the same network as SCL:
   #qMessage[1] := #s81_WtRFIDWriteOver;
END_REGION

REGION Network 55: Condition1 for STATE Num:82 Check RFID Write Retry Count Over
   RUNG wire#powerrail
      { S7_Templates := "SrcType := Int" } GT_Contact(in1 := #sRFWriteRetryCount, in2 := #iRetryCount)
      Coil( #c82_ChkWriteRetryCnt_T1 )
   END_RUNG
   // the same network as SCL:
   #c82_ChkWriteRetryCnt_T1 := #sRFWriteRetryCount > #iRetryCount;
END_REGION

REGION Network 56: Condition2 for STATE Num:82 Check RFID Write Retry Count Over
   RUNG wire#powerrail
      { S7_Templates := "SrcType := Int" } LE_Contact(in1 := #sRFWriteRetryCount, in2 := #iRetryCount)
      Coil( #c82_ChkWriteRetryCnt_T2 )
   END_RUNG
   // the same network as SCL:
   #c82_ChkWriteRetryCnt_T2 := #sRFWriteRetryCount <= #iRetryCount;
END_REGION

REGION Network 57: Transition for STATE Num:82 Check RFID Write Retry Count Over
   RUNG wire#powerrail
      Contact( #s82_ChkWriteRetryCnt )
      I_Contact( #sStWtResetRel )
      Contact( #sSst )
      wire#w1
      Contact( #c82_ChkWriteRetryCnt_T1 )
      Coil( #s82_ChkWriteRetryCnt_T1 )
   END_RUNG
   RUNG wire#w1
      I_Contact( #s82_ChkWriteRetryCnt_T1 )
      Contact( #c82_ChkWriteRetryCnt_T2 )
      Coil( #s82_ChkWriteRetryCnt_T2 )
   END_RUNG
   // the same network as SCL:
   #_w1 := #s82_ChkWriteRetryCnt AND NOT #sStWtResetRel AND #sSst;
   #s82_ChkWriteRetryCnt_T1 := #_w1 AND #c82_ChkWriteRetryCnt_T1;
   #s82_ChkWriteRetryCnt_T2 := #_w1 AND NOT #s82_ChkWriteRetryCnt_T1 AND #c82_ChkWriteRetryCnt_T2;
END_REGION

REGION Network 58: STATE Num:82 Check RFID Write Retry Count Over
   RUNG wire#powerrail
      Contact( #s82_ChkWriteRetryCnt )
      wire#w1
      I_Contact( #sStWtResetRel )
      I_Contact( #s82_ChkWriteRetryCnt_T1 )
      I_Contact( #s82_ChkWriteRetryCnt_T2 )
      wire#w2
      Coil( #s82_ChkWriteRetryCnt )
   END_RUNG
   RUNG wire#powerrail
      Contact( #s81_WtRFIDWriteOver_T1 )
   END_RUNG wire#w1
   RUNG wire#w2
      { S7_GenerateENO := "TRUE" } Move(in := 82, out1 => #StateNo)
   END_RUNG
   // the same network as SCL:
   #s82_ChkWriteRetryCnt := (#s82_ChkWriteRetryCnt OR #s81_WtRFIDWriteOver_T1) AND NOT #sStWtResetRel AND NOT #s82_ChkWriteRetryCnt_T1 AND NOT #s82_ChkWriteRetryCnt_T2;
   IF #s82_ChkWriteRetryCnt THEN #StateNo := 82; END_IF;
END_REGION

REGION Network 59: Actions for STATE Num:82 T1 - qError[3] := 1
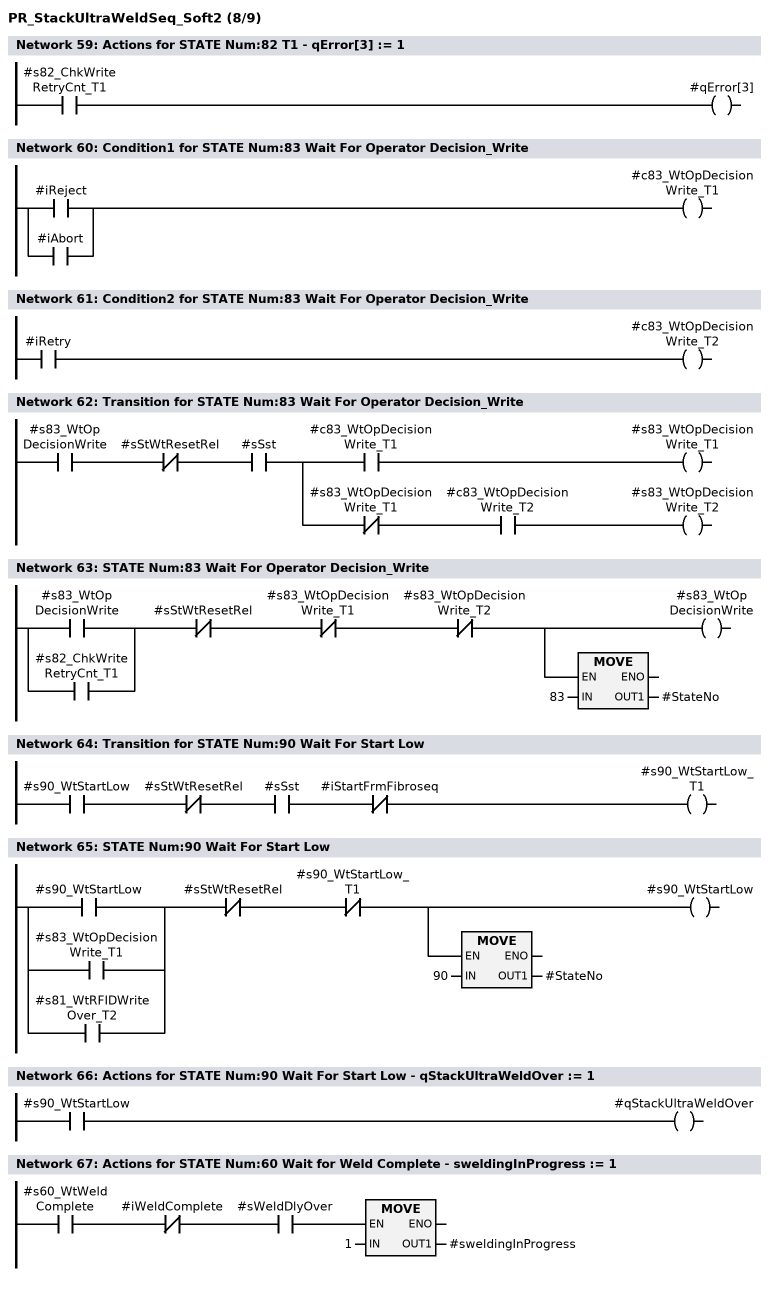
   RUNG wire#powerrail
      Contact( #s82_ChkWriteRetryCnt_T1 )
      Coil( #qError[3] )
   END_RUNG
   // the same network as SCL:
   #qError[3] := #s82_ChkWriteRetryCnt_T1;
END_REGION

REGION Network 60: Condition1 for STATE Num:83 Wait For Operator Decision_Write
   RUNG wire#powerrail
      Contact( #iReject )
      wire#w1
      Coil( #c83_WtOpDecisionWrite_T1 )
   END_RUNG
   RUNG wire#powerrail
      Contact( #iAbort )
   END_RUNG wire#w1
   // the same network as SCL:
   #c83_WtOpDecisionWrite_T1 := #iReject OR #iAbort;
END_REGION

REGION Network 61: Condition2 for STATE Num:83 Wait For Operator Decision_Write
   RUNG wire#powerrail
      Contact( #iRetry )
      Coil( #c83_WtOpDecisionWrite_T2 )
   END_RUNG
   // the same network as SCL:
   #c83_WtOpDecisionWrite_T2 := #iRetry;
END_REGION

REGION Network 62: Transition for STATE Num:83 Wait For Operator Decision_Write
   RUNG wire#powerrail
      Contact( #s83_WtOpDecisionWrite )
      I_Contact( #sStWtResetRel )
      Contact( #sSst )
      wire#w1
      Contact( #c83_WtOpDecisionWrite_T1 )
      Coil( #s83_WtOpDecisionWrite_T1 )
   END_RUNG
   RUNG wire#w1
      I_Contact( #s83_WtOpDecisionWrite_T1 )
      Contact( #c83_WtOpDecisionWrite_T2 )
      Coil( #s83_WtOpDecisionWrite_T2 )
   END_RUNG
   // the same network as SCL:
   #_w1 := #s83_WtOpDecisionWrite AND NOT #sStWtResetRel AND #sSst;
   #s83_WtOpDecisionWrite_T1 := #_w1 AND #c83_WtOpDecisionWrite_T1;
   #s83_WtOpDecisionWrite_T2 := #_w1 AND NOT #s83_WtOpDecisionWrite_T1 AND #c83_WtOpDecisionWrite_T2;
END_REGION

REGION Network 63: STATE Num:83 Wait For Operator Decision_Write
   RUNG wire#powerrail
      Contact( #s83_WtOpDecisionWrite )
      wire#w1
      I_Contact( #sStWtResetRel )
      I_Contact( #s83_WtOpDecisionWrite_T1 )
      I_Contact( #s83_WtOpDecisionWrite_T2 )
      wire#w2
      Coil( #s83_WtOpDecisionWrite )
   END_RUNG
   RUNG wire#powerrail
      Contact( #s82_ChkWriteRetryCnt_T1 )
   END_RUNG wire#w1
   RUNG wire#w2
      { S7_GenerateENO := "TRUE" } Move(in := 83, out1 => #StateNo)
   END_RUNG
   // the same network as SCL:
   #s83_WtOpDecisionWrite := (#s83_WtOpDecisionWrite OR #s82_ChkWriteRetryCnt_T1) AND NOT #sStWtResetRel AND NOT #s83_WtOpDecisionWrite_T1 AND NOT #s83_WtOpDecisionWrite_T2;
   IF #s83_WtOpDecisionWrite THEN #StateNo := 83; END_IF;
END_REGION

REGION Network 64: Transition for STATE Num:90 Wait For Start Low
   RUNG wire#powerrail
      Contact( #s90_WtStartLow )
      I_Contact( #sStWtResetRel )
      Contact( #sSst )
      I_Contact( #iStartFrmFibroseq )
      Coil( #s90_WtStartLow_T1 )
   END_RUNG
   // the same network as SCL:
   #s90_WtStartLow_T1 := #s90_WtStartLow AND NOT #sStWtResetRel AND #sSst AND NOT #iStartFrmFibroseq;
END_REGION

REGION Network 65: STATE Num:90 Wait For Start Low
   RUNG wire#powerrail
      Contact( #s90_WtStartLow )
      wire#w1
      I_Contact( #sStWtResetRel )
      I_Contact( #s90_WtStartLow_T1 )
      wire#w2
      Coil( #s90_WtStartLow )
   END_RUNG
   RUNG wire#powerrail
      Contact( #s83_WtOpDecisionWrite_T1 )
   END_RUNG wire#w1
   RUNG wire#powerrail
      Contact( #s81_WtRFIDWriteOver_T2 )
   END_RUNG wire#w1
   RUNG wire#w2
      { S7_GenerateENO := "TRUE" } Move(in := 90, out1 => #StateNo)
   END_RUNG
   // the same network as SCL:
   #s90_WtStartLow := (#s90_WtStartLow OR #s83_WtOpDecisionWrite_T1 OR #s81_WtRFIDWriteOver_T2) AND NOT #sStWtResetRel AND NOT #s90_WtStartLow_T1;
   IF #s90_WtStartLow THEN #StateNo := 90; END_IF;
END_REGION

REGION Network 66: Actions for STATE Num:90 Wait For Start Low - qStackUltraWeldOver := 1
   RUNG wire#powerrail
      Contact( #s90_WtStartLow )
      Coil( #qStackUltraWeldOver )
   END_RUNG
   // the same network as SCL:
   #qStackUltraWeldOver := #s90_WtStartLow;
END_REGION

REGION Network 67: Actions for STATE Num:60 Wait for Weld Complete - sweldingInProgress := 1
   RUNG wire#powerrail
      Contact( #s60_WtWeldComplete )
      I_Contact( #iWeldComplete )
      Contact( #sWeldDlyOver )
      { S7_GenerateENO := "TRUE" } Move(in := 1, out1 => #sweldingInProgress)
   END_RUNG
   // the same network as SCL:
   IF #s60_WtWeldComplete AND NOT #iWeldComplete AND #sWeldDlyOver THEN #sweldingInProgress := 1; END_IF;
END_REGION

REGION Network 68: Actions for STATE Num:80 Wait for Part Clamp Open - qFumeExtractorON := 0
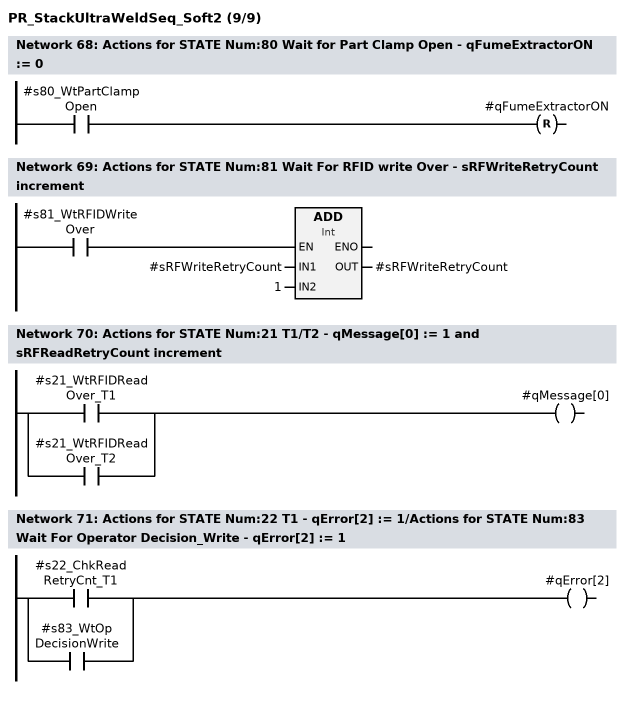
   RUNG wire#powerrail
      Contact( #s80_WtPartClampOpen )
      R_Coil( #qFumeExtractorON )
   END_RUNG
   // the same network as SCL:
   IF #s80_WtPartClampOpen THEN #qFumeExtractorON := FALSE; END_IF;
END_REGION

REGION Network 69: Actions for STATE Num:81 Wait For RFID write Over - sRFWriteRetryCount increment
   RUNG wire#powerrail
      Contact( #s81_WtRFIDWriteOver )
      { S7_Templates := "SrcType := Int"; S7_GenerateENO := "TRUE" } Add(in1 := #sRFWriteRetryCount, in2 := 1, out => #sRFWriteRetryCount)
   END_RUNG
   // the same network as SCL:
   IF #s81_WtRFIDWriteOver THEN #sRFWriteRetryCount := #sRFWriteRetryCount + 1; END_IF;
END_REGION

REGION Network 70: Actions for STATE Num:21 T1/T2 - qMessage[0] := 1 and sRFReadRetryCount increment
   RUNG wire#powerrail
      Contact( #s21_WtRFIDReadOver_T1 )
      wire#w1
      Coil( #qMessage[0] )
   END_RUNG
   RUNG wire#powerrail
      Contact( #s21_WtRFIDReadOver_T2 )
   END_RUNG wire#w1
   // the same network as SCL:
   #qMessage[0] := #s21_WtRFIDReadOver_T1 OR #s21_WtRFIDReadOver_T2;
END_REGION

REGION Network 71: Actions for STATE Num:22 T1 - qError[2] := 1/Actions for STATE Num:83 Wait For Operator Decision_Write - qError[2] := 1
   RUNG wire#powerrail
      Contact( #s22_ChkReadRetryCnt_T1 )
      wire#w1
      Coil( #qError[2] )
   END_RUNG
   RUNG wire#powerrail
      Contact( #s83_WtOpDecisionWrite )
   END_RUNG wire#w1
   // the same network as SCL:
   #qError[2] := #s22_ChkReadRetryCnt_T1 OR #s83_WtOpDecisionWrite;
END_REGION
END_FUNCTION_BLOCK
